{region 'Documentation'}
(*!
<summary>Checks held Abort cleanup and explicit completion without further enabled test work.</summary>
*)
{endregion}
FUNCTION_BLOCK Test_LifecycleAbort EXTENDS TestCaseLifecycleTestBase

SUPER^();

{region 'Documentation'}
(*!
<summary>Defines explicit exceptional-path stimuli and contract-derived observations.</summary>
*)
{endregion}
METHOD PROTECTED ConfigureScenario
FSubjectPreparationCount := 0;
FSubjectTestCount := 1;
FStepCount := 7;

{region "01 - Reset to Idle"}
// Establish Idle through the parent Reset request; both child results must be cleared.
FSteps[1].RequestReset := TRUE;
FSteps[1].ExpectedState := E_State.Idle;
FSteps[1].ExpectedResult := E_Result.NotEvaluated;
FSteps[1].ExpectedReady := TRUE;
FSteps[1].ExpectedPassedCount := 0;
FSteps[1].ExpectedFailedCount := 0;
FSteps[1].ExpectedHookCount := 6;
FSteps[1].ExpectedHooks[1].Hook := E_LifecycleHook.Reset;
FSteps[1].ExpectedHooks[1].State := E_State.Reset;
FSteps[1].ExpectedHooks[1].Enabled := TRUE;
FSteps[1].ExpectedHooks[2].Hook := E_LifecycleHook.Abort;
FSteps[1].ExpectedHooks[2].State := E_State.Idle;
FSteps[1].ExpectedHooks[2].Enabled := FALSE;
FSteps[1].ExpectedHooks[3].Hook := E_LifecycleHook.Preparations;
FSteps[1].ExpectedHooks[3].State := E_State.Idle;
FSteps[1].ExpectedHooks[3].Enabled := FALSE;
FSteps[1].ExpectedHooks[4].Hook := E_LifecycleHook.Tests;
FSteps[1].ExpectedHooks[4].State := E_State.Idle;
FSteps[1].ExpectedHooks[4].Enabled := FALSE;
FSteps[1].ExpectedHooks[5].Hook := E_LifecycleHook.Assertions;
FSteps[1].ExpectedHooks[5].State := E_State.Idle;
FSteps[1].ExpectedHooks[5].Enabled := FALSE;
FSteps[1].ExpectedHooks[6].Hook := E_LifecycleHook.Aggregate;
FSteps[1].ExpectedHooks[6].State := E_State.Idle;
FSteps[1].ExpectedHooks[6].Enabled := TRUE;
{endregion}

{region "02 - Accept Start"}
// Accept Start into Starting; processing and Assertion evaluation are not active yet.
FSteps[2].RequestStart := TRUE;
FSteps[2].ExpectedState := E_State.Starting;
FSteps[2].ExpectedResult := E_Result.NotEvaluated;
FSteps[2].ExpectedReady := FALSE;
FSteps[2].ExpectedPassedCount := 0;
FSteps[2].ExpectedFailedCount := 0;
FSteps[2].ExpectedHookCount := 5;
FSteps[2].ExpectedHooks[1].Hook := E_LifecycleHook.Abort;
FSteps[2].ExpectedHooks[1].State := E_State.Starting;
FSteps[2].ExpectedHooks[1].Enabled := FALSE;
FSteps[2].ExpectedHooks[2].Hook := E_LifecycleHook.Preparations;
FSteps[2].ExpectedHooks[2].State := E_State.Starting;
FSteps[2].ExpectedHooks[2].Enabled := FALSE;
FSteps[2].ExpectedHooks[3].Hook := E_LifecycleHook.Tests;
FSteps[2].ExpectedHooks[3].State := E_State.Starting;
FSteps[2].ExpectedHooks[3].Enabled := FALSE;
FSteps[2].ExpectedHooks[4].Hook := E_LifecycleHook.Assertions;
FSteps[2].ExpectedHooks[4].State := E_State.Starting;
FSteps[2].ExpectedHooks[4].Enabled := FALSE;
FSteps[2].ExpectedHooks[5].Hook := E_LifecycleHook.Aggregate;
FSteps[2].ExpectedHooks[5].State := E_State.Starting;
FSteps[2].ExpectedHooks[5].Enabled := TRUE;
{endregion}

{region "03 - Establish active execution"}
// Enter Running and evaluate both children; owner Result stays NotEvaluated until finalization.
FSteps[3].ExpectedState := E_State.Running;
FSteps[3].ExpectedResult := E_Result.NotEvaluated;
FSteps[3].ExpectedReady := FALSE;
FSteps[3].ExpectedPassedCount := 2;
FSteps[3].ExpectedFailedCount := 0;
FSteps[3].ExpectedHookCount := 5;
FSteps[3].ExpectedHooks[1].Hook := E_LifecycleHook.Abort;
FSteps[3].ExpectedHooks[1].State := E_State.Running;
FSteps[3].ExpectedHooks[1].Enabled := FALSE;
FSteps[3].ExpectedHooks[2].Hook := E_LifecycleHook.Preparations;
FSteps[3].ExpectedHooks[2].State := E_State.Running;
FSteps[3].ExpectedHooks[2].Enabled := FALSE;
FSteps[3].ExpectedHooks[3].Hook := E_LifecycleHook.Tests;
FSteps[3].ExpectedHooks[3].State := E_State.Running;
FSteps[3].ExpectedHooks[3].Enabled := TRUE;
FSteps[3].ExpectedHooks[4].Hook := E_LifecycleHook.Assertions;
FSteps[3].ExpectedHooks[4].State := E_State.Running;
FSteps[3].ExpectedHooks[4].Enabled := TRUE;
FSteps[3].ExpectedHooks[5].Hook := E_LifecycleHook.Aggregate;
FSteps[3].ExpectedHooks[5].State := E_State.Running;
FSteps[3].ExpectedHooks[5].Enabled := TRUE;
{endregion}

{region "04 - Request Abort and hold cleanup"}
// Request Abort and withhold cleanup completion; retain child results while entering Aborting.
FSteps[4].RequestAbort := TRUE;
FSteps[4].AbortCompleted := FALSE;
FSteps[4].ExpectedState := E_State.Aborting;
FSteps[4].ExpectedResult := E_Result.Abort;
FSteps[4].ExpectedReady := FALSE;
FSteps[4].ExpectedPassedCount := 2;
FSteps[4].ExpectedFailedCount := 0;
FSteps[4].ExpectedHookCount := 5;
FSteps[4].ExpectedHooks[1].Hook := E_LifecycleHook.Abort;
FSteps[4].ExpectedHooks[1].State := E_State.Aborting;
FSteps[4].ExpectedHooks[1].Enabled := TRUE;
FSteps[4].ExpectedHooks[2].Hook := E_LifecycleHook.Preparations;
FSteps[4].ExpectedHooks[2].State := E_State.Aborting;
FSteps[4].ExpectedHooks[2].Enabled := FALSE;
FSteps[4].ExpectedHooks[3].Hook := E_LifecycleHook.Tests;
FSteps[4].ExpectedHooks[3].State := E_State.Aborting;
FSteps[4].ExpectedHooks[3].Enabled := FALSE;
FSteps[4].ExpectedHooks[4].Hook := E_LifecycleHook.Assertions;
FSteps[4].ExpectedHooks[4].State := E_State.Aborting;
FSteps[4].ExpectedHooks[4].Enabled := FALSE;
FSteps[4].ExpectedHooks[5].Hook := E_LifecycleHook.Aggregate;
FSteps[4].ExpectedHooks[5].State := E_State.Aborting;
FSteps[4].ExpectedHooks[5].Enabled := TRUE;
{endregion}

{region "05 - Continue pending cleanup"}
// Continue active cleanup without a second Abort request; do not finalize before
// acknowledgement.
FSteps[5].AbortCompleted := FALSE;
FSteps[5].ExpectedState := E_State.Aborting;
FSteps[5].ExpectedResult := E_Result.Abort;
FSteps[5].ExpectedReady := FALSE;
FSteps[5].ExpectedPassedCount := 2;
FSteps[5].ExpectedFailedCount := 0;
FSteps[5].ExpectedHookCount := 5;
FSteps[5].ExpectedHooks[1].Hook := E_LifecycleHook.Abort;
FSteps[5].ExpectedHooks[1].State := E_State.Aborting;
FSteps[5].ExpectedHooks[1].Enabled := TRUE;
FSteps[5].ExpectedHooks[2].Hook := E_LifecycleHook.Preparations;
FSteps[5].ExpectedHooks[2].State := E_State.Aborting;
FSteps[5].ExpectedHooks[2].Enabled := FALSE;
FSteps[5].ExpectedHooks[3].Hook := E_LifecycleHook.Tests;
FSteps[5].ExpectedHooks[3].State := E_State.Aborting;
FSteps[5].ExpectedHooks[3].Enabled := FALSE;
FSteps[5].ExpectedHooks[4].Hook := E_LifecycleHook.Assertions;
FSteps[5].ExpectedHooks[4].State := E_State.Aborting;
FSteps[5].ExpectedHooks[4].Enabled := FALSE;
FSteps[5].ExpectedHooks[5].Hook := E_LifecycleHook.Aggregate;
FSteps[5].ExpectedHooks[5].State := E_State.Aborting;
FSteps[5].ExpectedHooks[5].Enabled := TRUE;
{endregion}

{region "06 - Acknowledge Abort cleanup"}
// Release AbortCompleted through its default TRUE value.
// The Abort hook enters Aborting, then all following hooks observe Completing.
FSteps[6].ExpectedState := E_State.Completing;
FSteps[6].ExpectedResult := E_Result.Abort;
FSteps[6].ExpectedReady := FALSE;
FSteps[6].ExpectedPassedCount := 2;
FSteps[6].ExpectedFailedCount := 0;
FSteps[6].ExpectedHookCount := 5;
FSteps[6].ExpectedHooks[1].Hook := E_LifecycleHook.Abort;
FSteps[6].ExpectedHooks[1].State := E_State.Aborting;
FSteps[6].ExpectedHooks[1].Enabled := TRUE;
FSteps[6].ExpectedHooks[2].Hook := E_LifecycleHook.Preparations;
FSteps[6].ExpectedHooks[2].State := E_State.Completing;
FSteps[6].ExpectedHooks[2].Enabled := FALSE;
FSteps[6].ExpectedHooks[3].Hook := E_LifecycleHook.Tests;
FSteps[6].ExpectedHooks[3].State := E_State.Completing;
FSteps[6].ExpectedHooks[3].Enabled := FALSE;
FSteps[6].ExpectedHooks[4].Hook := E_LifecycleHook.Assertions;
FSteps[6].ExpectedHooks[4].State := E_State.Completing;
FSteps[6].ExpectedHooks[4].Enabled := FALSE;
FSteps[6].ExpectedHooks[5].Hook := E_LifecycleHook.Aggregate;
FSteps[6].ExpectedHooks[5].State := E_State.Completing;
FSteps[6].ExpectedHooks[5].Enabled := TRUE;
{endregion}

{region "07 - Observe terminal Abort"}
// The following call reaches Completed; only aggregation remains in the recorded processing
// hooks.
FSteps[7].ExpectedState := E_State.Completed;
FSteps[7].ExpectedResult := E_Result.Abort;
FSteps[7].ExpectedReady := FALSE;
FSteps[7].ExpectedPassedCount := 2;
FSteps[7].ExpectedFailedCount := 0;
FSteps[7].ExpectedHookCount := 1;
FSteps[7].ExpectedHooks[1].Hook := E_LifecycleHook.Aggregate;
FSteps[7].ExpectedHooks[1].State := E_State.Completed;
FSteps[7].ExpectedHooks[1].Enabled := TRUE;
{endregion}
END_METHOD

END_FUNCTION_BLOCK

(* stored: Version 1.1.0.1
   POU Test_LifecycleAbort: Id {cd720fd3-2cab-46a4-befa-fa4baed24b3c}, SpecialFunc None
   Folder Internal: Id {078fc2ec-6094-405c-869d-49d72e592b5d}
   Method ConfigureScenario: Id {0c19af38-142a-4afb-970f-fc41ed8f691e} *)
